(* IEC 61131-3 sources: voltrus-explorers/apps/voltrus-plc/samples, 6 files *)

(* ---- BatchMixer.st ---- *)
PROGRAM BatchMixer
VAR
    (* State machine *)
    state : INT := 0;
    step_timer : INT := 0;

    (* Ingredient valves *)
    valve_a : BOOL := FALSE;
    valve_b : BOOL := FALSE;

    (* Process outputs *)
    mixer : BOOL := FALSE;
    heater : BOOL := FALSE;
    drain : BOOL := FALSE;

    (* Sensors *)
    level : REAL := 0.0;
    temperature : REAL := 20.0;

    (* Product *)
    batch_count : INT := 0;
    total_drained : REAL := 0.0;

    (* Recipe setpoints *)
    fill_level_a : REAL := 35.0;
    fill_level_b : REAL := 70.0;
    target_temp : REAL := 75.0;
    mix_time : INT := 150;
    drain_time : INT := 100;

    (* Alarms *)
    fault : BOOL := FALSE;
    fault_msg : INT := 0;

    (* Cycle counter *)
    cycles : DINT := 0;
END_VAR

    cycles := cycles + 1;
    step_timer := step_timer + 1;

    (* State machine *)
    IF state = 0 THEN
        (* IDLE *)
        valve_a := FALSE;
        valve_b := FALSE;
        mixer := FALSE;
        heater := FALSE;
        drain := FALSE;
        step_timer := 0;
        IF level <= 0.0 AND temperature < 30.0 THEN
            state := 1;
        END_IF;

    ELSIF state = 1 THEN
        (* FILL ingredient A *)
        valve_a := TRUE;
        IF level >= fill_level_a THEN
            valve_a := FALSE;
            state := 2;
            step_timer := 0;
        END_IF;

    ELSIF state = 2 THEN
        (* FILL ingredient B *)
        valve_b := TRUE;
        IF level >= fill_level_b THEN
            valve_b := FALSE;
            state := 3;
            step_timer := 0;
        END_IF;

    ELSIF state = 3 THEN
        (* HEAT to target *)
        mixer := TRUE;
        heater := TRUE;
        IF temperature >= target_temp THEN
            heater := FALSE;
            state := 4;
            step_timer := 0;
        END_IF;

    ELSIF state = 4 THEN
        (* MIX for duration *)
        mixer := TRUE;
        IF step_timer >= mix_time THEN
            mixer := FALSE;
            state := 5;
            step_timer := 0;
        END_IF;

    ELSIF state = 5 THEN
        (* DRAIN product *)
        drain := TRUE;
        IF step_timer >= drain_time THEN
            drain := FALSE;
            batch_count := batch_count + 1;
            state := 0;
            step_timer := 0;
        END_IF;

    END_IF;

    (* Watchdog: fault if any state takes too long *)
    IF step_timer > 500 THEN
        fault := TRUE;
        fault_msg := state;
    END_IF;

    (* Simulate process dynamics *)
    IF valve_a THEN
        level := level + 0.8;
    END_IF;
    IF valve_b THEN
        level := level + 1.0;
    END_IF;
    IF drain THEN
        level := level - 1.2;
        total_drained := total_drained + 1.2;
    END_IF;
    IF heater THEN
        temperature := temperature + 0.4;
    END_IF;
    IF mixer AND NOT heater THEN
        temperature := temperature - 0.08;
    END_IF;

    (* Clamp *)
    IF level > 100.0 THEN
        level := 100.0;
    END_IF;
    IF level < 0.0 THEN
        level := 0.0;
    END_IF;
    IF temperature < 0.0 THEN
        temperature := 0.0;
    END_IF;
    IF temperature > 120.0 THEN
        temperature := 120.0;
    END_IF;

END_PROGRAM

(* ---- Counter.st ---- *)
PROGRAM Counter
VAR
    counter : INT := 0;
    max_count : INT := 100;
    done : BOOL := FALSE;
    cycles : DINT := 0;
    direction : INT := 1;
END_VAR

    cycles := cycles + 1;

    counter := counter + direction;

    IF counter >= max_count THEN
        direction := -1;
        done := TRUE;
    ELSIF counter <= 0 THEN
        direction := 1;
        done := FALSE;
    END_IF;

END_PROGRAM

(* ---- ESP32_Tester.st ---- *)
PROGRAM ESP32_Tester
VAR
    (* Inputs from ESP32 — mapped to Modbus holding registers *)
    counter : DINT;        (* Reg 0: auto-incrementing counter, 1s interval *)
    random_val : DINT;     (* Reg 1: random value 0-999 *)

    (* Outputs to ESP32 — mapped to Modbus holding registers *)
    buzzer : BOOL := FALSE;     (* Reg 10: buzzer on/off *)
    red : DINT := 0;            (* Reg 11: RGB red 0-255 *)
    green : DINT := 0;          (* Reg 12: RGB green 0-255 *)
    blue : DINT := 0;           (* Reg 13: RGB blue 0-255 *)

    (* Relay outputs — mapped to Modbus coils 0-5 *)
    relay0 : BOOL := FALSE;
    relay1 : BOOL := FALSE;
    relay2 : BOOL := FALSE;
    relay3 : BOOL := FALSE;
    relay4 : BOOL := FALSE;
    relay5 : BOOL := FALSE;

    (* Internal logic *)
    cycle : DINT := 0;
    phase : DINT := 0;
    step_timer : TON;
    flash_timer : TON;
END_VAR

    cycle := cycle + 1;

    (* Step timer: advance phase every 2 seconds *)
    step_timer(IN := TRUE, PT := T#2S);
    IF step_timer.Q THEN
        step_timer(IN := FALSE, PT := T#0MS);
        phase := phase + 1;
        IF phase > 5 THEN
            phase := 0;
        END_IF;
    END_IF;

    (* Flash timer for visual feedback *)
    flash_timer(IN := TRUE, PT := T#500MS);
    IF flash_timer.Q THEN
        flash_timer(IN := FALSE, PT := T#0MS);
    END_IF;

    (* Buzzer: beep when counter is in upper half *)
    IF counter > 500 THEN
        buzzer := TRUE;
    ELSE
        buzzer := FALSE;
    END_IF;

    (* Relay pattern based on phase *)
    CASE phase OF
        0:  (* All off *)
            relay0 := FALSE; relay1 := FALSE; relay2 := FALSE;
            relay3 := FALSE; relay4 := FALSE; relay5 := FALSE;
        1:  (* Chase right *)
            relay0 := TRUE; relay1 := FALSE; relay2 := FALSE;
            relay3 := FALSE; relay4 := FALSE; relay5 := FALSE;
        2:  (* Chase right *)
            relay0 := FALSE; relay1 := TRUE; relay2 := FALSE;
            relay3 := FALSE; relay4 := FALSE; relay5 := FALSE;
        3:  (* Chase right *)
            relay0 := FALSE; relay1 := FALSE; relay2 := TRUE;
            relay3 := FALSE; relay4 := FALSE; relay5 := FALSE;
        4:  (* Chase right *)
            relay0 := FALSE; relay1 := FALSE; relay2 := FALSE;
            relay3 := TRUE; relay4 := FALSE; relay5 := FALSE;
        5:  (* All on *)
            relay0 := TRUE; relay1 := TRUE; relay2 := TRUE;
            relay3 := TRUE; relay4 := TRUE; relay5 := TRUE;
    END_CASE;

    (* RGB LED: cycle through colors based on phase *)
    CASE phase OF
        0:  red := 255; green := 0;   blue := 0;     (* Red *)
        1:  red := 0;   green := 255; blue := 0;     (* Green *)
        2:  red := 0;   green := 0;   blue := 255;   (* Blue *)
        3:  red := 255; green := 255; blue := 0;     (* Yellow *)
        4:  red := 255; green := 0;   blue := 255;   (* Magenta *)
        5:  red := 0;   green := 255; blue := 255;   (* Cyan *)
    END_CASE;

END_PROGRAM

(* ---- MotorControl.st ---- *)
PROGRAM MotorControl
VAR
    (* Inputs *)
    start_btn : BOOL := FALSE;
    stop_btn : BOOL := FALSE;
    emergency_stop : BOOL := FALSE;
    overload_trip : BOOL := FALSE;

    (* Outputs *)
    motor_running : BOOL := FALSE;
    fault : BOOL := FALSE;
    speed : INT := 0;
    fault_code : INT := 0;

    (* Parameters *)
    target_speed : INT := 1000;
    ramp_rate : INT := 10;
    decel_rate : INT := 25;

    (* Runtime *)
    run_time : DINT := 0;
    start_delay : INT := 0;
END_VAR

    run_time := run_time + 1;

    (* Safety: check overload *)
    IF overload_trip THEN
        fault := TRUE;
        fault_code := 1;
        motor_running := FALSE;
    END_IF;

    (* Safety: emergency stop *)
    IF emergency_stop THEN
        fault := TRUE;
        fault_code := 2;
        motor_running := FALSE;
    END_IF;

    (* Start logic: latch on *)
    IF start_btn AND NOT stop_btn AND NOT fault THEN
        IF (NOT motor_running) AND (speed = 0) THEN
            start_delay := start_delay + 1;
            IF start_delay > 10 THEN
                motor_running := TRUE;
                start_delay := 0;
            END_IF;
        ELSE
            motor_running := TRUE;
            start_delay := 0;
        END_IF;
    END_IF;

    (* Stop logic *)
    IF stop_btn THEN
        motor_running := FALSE;
        start_delay := 0;
    END_IF;

    (* Fault reset: hold stop for 2 seconds *)
    IF stop_btn AND fault THEN
        start_delay := start_delay + 1;
        IF start_delay > 20 THEN
            fault := FALSE;
            fault_code := 0;
            start_delay := 0;
        END_IF;
    END_IF;

    (* Speed ramping *)
    IF motor_running THEN
        IF speed < target_speed THEN
            speed := speed + ramp_rate;
            IF speed > target_speed THEN
                speed := target_speed;
            END_IF;
        END_IF;
    ELSE
        IF speed > 0 THEN
            speed := speed - decel_rate;
            IF speed < 0 THEN
                speed := 0;
            END_IF;
        END_IF;
    END_IF;

END_PROGRAM

(* ---- TankLevel.st ---- *)
PROGRAM TankLevel
VAR
    (* Process variable *)
    level : REAL := 25.0;
    temperature : REAL := 20.0;

    (* Setpoints *)
    level_setpoint : REAL := 50.0;
    temp_setpoint : REAL := 65.0;
    deadband : REAL := 3.0;

    (* Outputs *)
    inlet_valve : BOOL := FALSE;
    outlet_valve : BOOL := FALSE;
    heater : BOOL := FALSE;
    cooling_valve : BOOL := FALSE;

    (* Alarms *)
    high_level_alarm : BOOL := FALSE;
    low_level_alarm : BOOL := FALSE;
    high_temp_alarm : BOOL := FALSE;

    (* Simulation parameters *)
    inlet_flow : REAL := 1.0;
    outlet_flow : REAL := 0.6;
    heat_rate : REAL := 0.3;
    cool_rate : REAL := 0.15;
    ambient_loss : REAL := 0.05;

    (* Statistics *)
    cycles : DINT := 0;
    total_inlet_time : DINT := 0;
    total_outlet_time : DINT := 0;
END_VAR

    cycles := cycles + 1;

    (* Level control - bang-bang with deadband *)
    IF level < level_setpoint - deadband THEN
        inlet_valve := TRUE;
        outlet_valve := FALSE;
    ELSIF level > level_setpoint + deadband THEN
        inlet_valve := FALSE;
        outlet_valve := TRUE;
    END_IF;

    (* Temperature control *)
    IF temperature < temp_setpoint - deadband THEN
        heater := TRUE;
        cooling_valve := FALSE;
    ELSIF temperature > temp_setpoint + deadband THEN
        heater := FALSE;
        cooling_valve := TRUE;
    END_IF;

    (* Alarms *)
    high_level_alarm := level > 90.0;
    low_level_alarm := level < 10.0;
    high_temp_alarm := temperature > 85.0;

    (* Emergency shutdown *)
    IF high_level_alarm THEN
        inlet_valve := FALSE;
    END_IF;
    IF high_temp_alarm THEN
        heater := FALSE;
    END_IF;

    (* Simulate process dynamics *)
    IF inlet_valve THEN
        level := level + inlet_flow;
        total_inlet_time := total_inlet_time + 1;
    END_IF;
    IF outlet_valve THEN
        level := level - outlet_flow;
        total_outlet_time := total_outlet_time + 1;
    END_IF;
    IF heater THEN
        temperature := temperature + heat_rate;
    END_IF;
    IF cooling_valve THEN
        temperature := temperature - cool_rate;
    END_IF;

    (* Ambient heat loss *)
    temperature := temperature - ambient_loss;

    (* Clamp values *)
    IF level > 100.0 THEN
        level := 100.0;
    END_IF;
    IF level < 0.0 THEN
        level := 0.0;
    END_IF;
    IF temperature < 0.0 THEN
        temperature := 0.0;
    END_IF;
    IF temperature > 100.0 THEN
        temperature := 100.0;
    END_IF;

END_PROGRAM

(* ---- TrafficLight.st ---- *)
PROGRAM TrafficLight
VAR
    state : INT := 0;
    timer : INT := 0;
    red : BOOL := TRUE;
    yellow : BOOL := FALSE;
    green : BOOL := FALSE;
    flash : BOOL := FALSE;
    flash_counter : INT := 0;
    pedestrian_waiting : BOOL := FALSE;
END_VAR

    timer := timer + 1;
    flash_counter := flash_counter + 1;
    flash := (flash_counter MOD 20) > 10;

    IF state = 0 THEN
        (* Red - stop traffic *)
        red := TRUE;
        yellow := FALSE;
        green := FALSE;
        IF timer > 100 THEN
            state := 1;
            timer := 0;
        END_IF;

    ELSIF state = 1 THEN
        (* Red + Yellow - prepare to go *)
        red := TRUE;
        yellow := TRUE;
        green := FALSE;
        IF timer > 30 THEN
            state := 2;
            timer := 0;
        END_IF;

    ELSIF state = 2 THEN
        (* Green - go *)
        red := FALSE;
        yellow := FALSE;
        green := TRUE;
        IF timer > 100 THEN
            state := 3;
            timer := 0;
        END_IF;

    ELSIF state = 3 THEN
        (* Yellow - warning *)
        red := FALSE;
        yellow := TRUE;
        green := FALSE;
        IF timer > 40 THEN
            state := 0;
            timer := 0;
        END_IF;
    END_IF;

END_PROGRAM
